(* IEC 61131-3 sources: Masterarbeit/sigmatek/lasalclass2/PW022_virtualization/Network/HW_Network, 1 file *)

(* ---- ONE_HW_Network_Table.st ---- *)
#define OBJECTS_CONFIG

//Define part of class Varan_Base
#ifndef _T_VARANBASE_H
#define _T_VARANBASE_H

#define	VARAN_PLL_OFFSET		16#0140
#define VARAN_MULTIPLE_OFFSET	16#01AC

// version of serial number validation (16#10 = 1.0)
#define SERNO_VALIDATION_VERSION 16#10

#define IsTransparent_IS_AVAILABLE

// Defines for Mutex Generation
#define VARAN_STR_MUTEX_NAME_SEPERATOR ".."
#define VARAN_MUTEX_NAME_END_LENGTH 5
#define VARAN_MUTEX_NAME_MAX_LENGTH 32

#define VARAN_SPI_IDENT_LICENCENO_OFFSET    16#14
#define VARAN_SPI_IDENT_HARDWAREVER_OFFSET  16#18

#endif // _T_VARANBASE_H
#include "..\..\Class\HwControl\HwControl.h"
#include "..\..\Source\interfaces\lsl_st_hardwaretree.h"
//Define part of class BusInterfaceVARAN
#define BUSIF_VARAN_MAX_NR_DO     100
#define BUSIF_VARAN_MAX_NR_MOVEDO 100

#define BUSIF_VARAN_MAX_SDO 1

#define BUSIF_VARAN_BUS_READY_VER 16#1109
#include "..\..\Source\BusInterface.h"
#include "..\..\Source\interfaces\lsl_st_mt.h"
#include "..\..\Source\interfaces\lsl_st_pci.h"
#include "..\..\Class\HwControl\watchdog.h"
#include "..\..\Source\interfaces\lsl_st_sysinfo.h"
#include "..\..\Source\interfaces\lsl_st_systrace.h"
#include "..\..\Class\HwControl\_HWKScope.h"
#include <.\lsl_st_mt.h>
//Define part of class SdiasBase
//Address to access the Dataobject list via SPI SDO Read
#define SDIAS_SPI_DATA_OBJECT_LIST_PAGE_ADDRESS               16#FFFF
#define SDIAS_SPI_DATA_OBJECT_LIST_PAGE_OFFSET                16#00
#define SDIAS_SPI_DATA_OBJECT_LIST_IDENTIFIER                 16#12345678

//Defines the number of optional list elements in the SPI List

#define SDIAS_SPI_NUMBER_OF_OPTIONAL_ELEMENTS                 16

#define SDIAS_SPI_HEADER_BEFORE_OPTIONAL_ELEMENTS             16#18
#define SDIAS_SPI_HARDWARE_VERSION_OFFSET                     16#C
#define SDIAS_SPI_VENDOR_ID_OFFSET                            16#0

#define SDIAS_SPI_MASTER_ADRESS_TRANSMIT_BUFFER0              16#0000
#define SDIAS_SPI_MASTER_ADRESS_TRANSMIT_BUFFER1              16#0080
#define SDIAS_SPI_MASTER_ADRESS_RECEIVE_BUFFER0               16#0000
#define SDIAS_SPI_MASTER_ADRESS_RECEIVE_BUFFER1               16#0080
#define SDIAS_SPI_MASTER_ADRESS_PAGE_ADRESS                   16#0100
#define SDIAS_SPI_MASTER_ADRESS_PREDEFINED_COMMAND_REGISTER   16#0102
#define SDIAS_SPI_MASTER_ADRESS_SINGLE_COMMAND_REGISTER       16#0103
#define SDIAS_SPI_MASTER_ADRESS_STATUS_REGISTER               16#0104
#define SDIAS_SPI_MASTER_ADRESS_REQUEST_REGISTER              16#0105
#define SDIAS_SPI_MASTER_ADRESS_GRANT_REGISTER                16#0106
#define SDIAS_SPI_MASTER_ADRESS_CLEAR_REQUEST_REGISTER        16#0107
#define SDIAS_SPI_MASTER_ADRESS_FEATURE_REGISTER              16#0108

#define SDIAS_SPI_MASTER_SOFTWARE_REQUEST                     1

#define SDIAS_SPI_MASTER_COMMAND_PAGE_READ                    16#01
#define SDIAS_SPI_MASTER_COMMAND_PAGE_PROGRAM                 16#02
#define SDIAS_SPI_MASTER_COMMAND_SECTOR_ERASE                 16#03
#define SDIAS_SPI_MASTER_COMMAND_REBOOT_FPGA                  16#F0

#define SDIAS_SPI_MASTER_STATE_BUSY                           16#00
#define SDIAS_SPI_MASTER_STATE_READY                          16#01

#define SDIAS_SPI_SECTOR_SIZE                                 65536 // 256*256
#define SDIAS_SPI_PAGE_SIZE                                   256

#define SDIAS_SPI_WRITE_MAX_RETRIES                           2
#define SDIAS_SPI_TIMEOUT                                     500  //timeout for spi accesses
#define SDIAS_SPI_LOCK_TIMEOUT                                6   //this value is multiplied with the buscycletime [µs] (6*1000=6.000 msec timeout)

//SPI List IDs
#define SDIAS_SPI_IDENTIFICATION_LIST_ID  1
#define SDIAS_SPI_FLASH_CONFIGURATION_ID  2
#define SDIAS_SPI_VENDOR_NAME_ID          3
#define SDIAS_SPI_DEVICE_NAME_ID          4
#define SDIAS_SPI_SERIAL_NUMBER_ID        5
#define SDIAS_SPI_ORDERING_NUMBER_ID      6
#define SDIAS_SPI_DOCUMENTATION_PDF_ID    7
#define SDIAS_SPI_CALIB_DATA_ID           10
#define SDIAS_SPI_PDO_INFORMATION_ID      128

//SPI Access
#define SDIAS_SPI_ACCESS_ID_HW_TREE          1
#define SDIAS_SPI_ACCESS_ID_HWK_INTERNAL     2
#include "..\..\Class\SdiasManager\SdiasManager.h"
#include "..\..\Class\SdiasBase\SdiasBase.h"
//Define part of class PW022
#define DEVICE_ID_PW022                     1089
// address offsets for SDO communication
#define PW022_ADDR_CFG_MODUL                16#004
// timeouts
#define PW022_SDO_RESPONSE_TIMEOUT          SDIAS_SDO_TIMEOUT * 2
#define PW022_MIN_PERIODE_TIME              100  //minimal allowed periode time * 500nsec
#define PW022_MAX_PERCENT                 10000  //maximal value for percent (100.00)
//Define part of class SafetyUDP
#define SAFETY_UDP_MAX_SOCKETS                6     // Max number of socket

#define SAFETY_UDP_CLT_SEND_OK                0    // Send ok
#define SAFETY_UDP_CLT_INVALID_HANDLE        -1    // Invalid handle
#define SAFETY_UDP_CLT_NOT_OPEN              -2    // Socket is not open
#define SAFETY_UDP_CLT_SEND_FAILED           -3    // Send failed
#define SAFETY_UDP_CLT_SEND_BUFFER_FULL      -4    // Send buffer is full
#define SAFETY_UDP_CLT_DATA_TO_BIG           -5    // Data to big

#define SAFETY_UDP_MAXIMUM_SEGMENT_SIZE    1452    // Maximum of user data

#define SAFETY_UDP_TIMEOUT_OPENSOCKET    (1000)    //timeout for opening socket

#define SAFETY_UDP_RECEIVE_TIMEOUT          800

#define SAFETY_UDP_TX_BUFFER_SIZE          1024
//Define part of class SafetyManager
#define LogBufferSize 1000
#include "..\..\Class\SafetyManager\SafetyManager.h"
#include "..\..\Source\interfaces\lsl_st_safetydll.h"
//Define part of class SdiasManager
#define SDIAS_SDO_MAX_LENGTH              128
#define SDIAS_SDO_RINGBUFFER_NO            64
#define SDIAS_SDO_CHANNEL_NO                3   // fixed in the VI hardware to be 3

// watchdog trigger interval (after 130ms of no trigger the SDIAS HW goes into reset again and takes at least another 10ms to be ready again)
#define SDIAS_WATCHDOG_TRIGGER_TIME        40

// time needed by sdias modules to start up after the watchdog is triggered the first time in ms
#define SDIAS_HARDWARE_STARTUP_TIME        15

// sdias manager needs 2 ticks to handle event for read task (measure sync time)
#define SDIAS_SYNC_MEASURE_TICKS            2

// after activating the PLL SyncOut it takes 3 cycles until the SDIAS sync can be injected
#define SDIAS_CYCLES_WAIT_AFTER_SYNC_ENABLE 3

// wait 1 bus cycle at start to get valid numbers in the task info
#define SDIAS_TASKINFO_READY_TICKS          1

// time to wait (in ms) until other tasks in the same or lower priority than post init have done their stuff
#define SDIAS_WAIT_TIME_IN_POST_INIT        1

#define SIZE_PER_SDIAS_CLIENT               16#0400

// for far memory accesses: 1 module can hold maximum 256 1K blocks (0-255)
#define SDIAS_1K_BLOCK_NO                       256

// far memory accesses maximum length in bytes
#define SDIAS_MAX_SIZE_FAR_MEM_ACCESS           127

#define SDIAS_OFFSET_HW_CONFIG              16#FF00
#define SDIAS_OFFSET_TASK_EVENT_IDS         16#FF10
#define SDIAS_OFFSET_FEATURE_INFO           16#FF18
#define SDIAS_OFFSET_APPLI_LED_STATES       16#FF20
#define SDIAS_OFFSET_SYNC_INJECTION_CFG     16#FF3D
#define SDIAS_OFFSET_TRIGGER_UNIT_SETUP_0   16#FF41
#define SDIAS_OFFSET_TRIGGER_UNIT_SETUP_1   16#FF45
#define SDIAS_OFFSET_TASK_START_CFG_0       16#FF60
#define SDIAS_OFFSET_TASK_CONFIG_0          16#FF86
#define SDIAS_OFFSET_TASK_CONFIG_1          16#FF96
#define SDIAS_OFFSET_TASK_INFO_1            16#FF94
#define SDIAS_OFFSET_TASK_HANDSHAKE_1       16#FF9B
#define SDIAS_OFFSET_TASK_DURATION_TIME_1   16#FF9C
#define SDIAS_OFFSET_TASK_DURATION_TIME_2   16#FFAC
#define SDIAS_OFFSET_TASK_CONFIG_2          16#FFA6

#define SDIAS_RETRIES_ALLOWED         2

// mask to get global error flag out of message counter byte of SDO responses
#define SDIAS_MASK_GLOBAL_ERROR_FLAG        16#80

// mask to get message counter out of message counter byte of SDO responses
#define SDIAS_MASK_MESSAGE_COUNTER          16#3F

#define SDIAS_EVENT_MASK_ID_SYNC_OUT0       16#10
#define SDIAS_EVENT_MASK_ID_SYNC_OUT1       16#11
#define SDIAS_EVENT_MASK_ID_SYNC_OUT2       16#12
#define SDIAS_EVENT_MASK_ID_SYNC_OUT3       16#13

#define SDIAS_MANAGER_SYNC_SYNCOUT_ID       16#85
#define SDIAS_TASK_START_EVENT_SYNCOUT_ID   16#86

#define SDIAS_PLACE_NO_MODULE_ADDED_SO_FAR  16#80000000

#define SDIAS_TRIGGER_UNIT_BYTE_SIZE        2

#define SDIAS_WAIT_TIME_FIRMWARE_HANDSHAKE  5 * 1000

// if the firmware version is below this, there might be problems with SCP111 and other modules => print warning at startup
#define SDIAS_FW_VERSION_SDO_ERROR_FIXED    16#120

// if the protocol version ist below this, Control Read/Broadcast Write Command is not supported by sdiasmanager
#define SDIAS_PROTOCOLVERSION_BROADCAST     16#120

// if the cil version ist below this, Control Read/Broadcast Write Command is not supported by OS for local SDIAS.
#define SDIAS_CILVERSION_BROADCAST         16#5001

// timeout for blocking the init during initialisation (in ms)
#define SDIAS_INIT_BLOCK_TIMEOUT            20 * 1000

#define SDIAS_MUTEX_NAME_END_LENGTH 3
#define SDIAS_MUTEX_NAME_MAX_LENGTH 32
#define SDIAS_MUTEX_STR_SEPERATOR   ".."

//#define SDIAS_RT_TIME_MEASUREMENT
#ifdef SDIAS_RT_TIME_MEASUREMENT
  #pragma message("ATTENTION: SDIAS real time measurement is active and needs additional ressources in the realtime task")
#endif

(* SDIAS data object commands  *)
#define	 SDIAS_CMD_END							  0x00			(* End command										          *)
#define	 SDIAS_CMD_ACC_MEMORY				  0x01			(* Access dpram memory								      *)
#define	 SDIAS_CMD_ACC_CONTROL				0x02			(* Access dpram control memory						  *)
#define	 SDIAS_CMD_GLOBAL						  0x03			(* SDIAS global command								      *)
#define	 SDIAS_CMD_COPY_LOCAL					0x04			(* DPRAM copy command in local dpram				*)
#define	 SDIAS_CMD_JMP_LOCAL					0x05			(* DPRAM jump command in local dpram 				*)
#define  SDIAS_CMD_ACC_MEMORY_FAR     0x07      (* SDIAS Far Memory Access                  *)

(* SDIAS defines for data object handling *)
// Write data oject list
#define	 SDIAS_DOL_WRITE_USAGE_DOL_EMPTY	  0x20			(* Usage of empty write dol list (wachtdog trigger + end command)   *)
#define	 SDIAS_DOL_WRITE_USAGE_DTA_EMPTY	  0x03			(* Usage of empty write dol data (DO ctrl of 2x copy command for task information + DO ctrl of watchdog trigger      *)
#define	 SDIAS_DOL_WRITE_OFFSET_END_CMD			0x10			(* One data object in list - offset = 1 DO size = 0x10						  *)
#define	 SDIAS_DOL_WRITE_OFFSET_FIRST_DTA		0x02			(* Offset of first data byte of second copy command = 2 (DO ctrl)   *)
#define	 SDIAS_DOL_WRITE_OFFSET_LAST_DTA		0x02			(* Offset of last data byte of second copy command = 2 (DO ctrl )   *)

// Read data oject list
#define	 SDIAS_DOL_READ_USAGE_DOL_EMPTY	    0x30			(* Usage of empty read dol list (2x task info copy command + end command)   *)
#define	 SDIAS_DOL_READ_USAGE_DTA_EMPTY	    0x0D			(* Usage of empty write dol data (DO ctrl of 2x copy command for task information + DO ctrl of watchdog trigger      *)
#define	 SDIAS_DOL_READ_OFFSET_END_CMD			0x20			(* One data object in list - offset = 1 DO size = 0x10						          *)
#define	 SDIAS_DOL_READ_OFFSET_FIRST_DTA		0x07			(* Offset of first data byte of second copy command = 7 = DO state          *)
#define	 SDIAS_DOL_READ_OFFSET_LAST_DTA		  0x0C			(* Offset of last data byte of second copy command = 12 (last byte of task information)       *)

//Versionsnumber where SDIAS SPI Read Accesses are available
#define  SDIAS_SDO_SPI_FIRMWARE_VERSION_AVAILABLE 16#0120

//error info mask
#define  SDIAS_ERROR_INFO_MASK    2#1000011000011111

// Broadcast DO Info
#define SDIAS_OFFSET_CLIENT_CTRLTIMESTAMP   16#0190
#define SDIAS_NR_TIMEBROADCAST_DOS 2
#define SDIAS_TIMEBROADCAST_SUBCMD 16#B0
#include "..\..\source\interfaces\lsl_st_pll.h"
//Define part of class VaranManager
#define SIZE_PAYLOAD_FRAME_HEADER_DO      16#38  // Const because datasize is in the Payload DOs
#define SIZE_PAYLOAD_IRQ_FRAME_HEADER_DO  16#40  // Const because datasize is in the Payload DOs

#define VM_MAX_POST_INIT_MODULES  1000

#define VM_OBJECT_PATH            16#81000002   // Object Path for Varanmanager Length = 2 (First 2byte), Domain = 0 (3rd byte), Escape Sequence Varan (4th byte)
#include "..\..\Class\VaranManager\VaranManager.h"
#include "..\..\Source\interfaces\lsl_st_kernel.h"
//Define part of class VaranManager_2
// needed to use the same code as the other managing modules
#define VM2_SYNCHRON SuperiorSystemOK

#define VM2_SDO_INIT_CMD_LENGTH   12
//Define part of class VI021
#define DEVICE_ID_VI022 1233

FUNCTION GLOBAL TAB ONE_HW_Network
-1$UINT, 0$UINT,
0$UINT, 0$UINT,

26$UDINT,
TO_UDINT(2897291062), "ASCII_BIN", 1$UINT, 21$UINT, 1$UINT,
TO_UDINT(24783181), "BusInterfaceVARAN", 1$UINT, 75$UINT, 0$UINT,
TO_UDINT(794617671), "CriticalSection", 0$UINT, 4$UINT, 2$UINT,
TO_UDINT(3238133653), "Hub_Base", 1$UINT, 21$UINT, 1$UINT,
TO_UDINT(1770276445), "Hub_Base_Root", 2$UINT, 11$UINT, 2$UINT,
TO_UDINT(3078259981), "HwcLogging", 1$UINT, 0$UINT, 1$UINT,
TO_UDINT(2471641665), "HwControl", 5$UINT, 21$UINT, 1$UINT,
TO_UDINT(1193052171), "HwControlBase", 1$UINT, 10$UINT, 0$UINT,
TO_UDINT(4260294091), "HWRtPostScan", 1$UINT, 0$UINT, 1$UINT,
TO_UDINT(2225119864), "MerkerEx", 1$UINT, 22$UINT, 4$UINT,
TO_UDINT(2837966764), "PW022", 1$UINT, 5$UINT, 3$UINT,
TO_UDINT(3591333481), "RamFile", 1$UINT, 9$UINT, 1$UINT,
TO_UDINT(1799751072), "SafetyManager", 2$UINT, 26$UINT, 1$UINT,
TO_UDINT(3727715967), "SafetyUDP", 1$UINT, 4$UINT, 0$UINT,
TO_UDINT(3175101883), "SdiasBase", 1$UINT, 60$UINT, 0$UINT,
TO_UDINT(4173303375), "SdiasHubBase", 1$UINT, 10$UINT, 1$UINT,
TO_UDINT(2118381352), "SdiasManager", 1$UINT, 97$UINT, 1$UINT,
TO_UDINT(736632136), "Steuerung", 0$UINT, 0$UINT, 1$UINT,
TO_UDINT(1850111279), "String", 1$UINT, 11$UINT, 4$UINT,
TO_UDINT(2898603620), "StringInternal", 1$UINT, 85$UINT, 0$UINT,
TO_UDINT(862125188), "Varan_Base", 2$UINT, 20$UINT, 0$UINT,
TO_UDINT(2940693151), "VaranManager", 3$UINT, 7$UINT, 0$UINT,
TO_UDINT(4019434288), "VaranManager_2", 2$UINT, 9$UINT, 1$UINT,
TO_UDINT(4035182347), "VaranManager_Base", 1$UINT, 26$UINT, 0$UINT,
TO_UDINT(262695706), "VI021", 1$UINT, 101$UINT, 1$UINT,
TO_UDINT(3232495061), "VirtualBaseInit", 1$UINT, 3$UINT, 0$UINT,

1$UINT, TO_UDINT(1973273396), "VARANMANAGER_21\_BASE\ASCII_BIN1",

1$UINT, TO_UDINT(2972590922), "HWCONTROL1\SAFETYMANAGER\UDPRECEIVEDATA",
1$UINT, TO_UDINT(1868223583), "HWCONTROL1\SAFETYMANAGER\UDPSENDDATA",

1$UINT, TO_UDINT(658018123), "VI0211\HUB_BASE1",

1$UINT, TO_UDINT(980975553), "VARANMANAGER_21\HUB_BASE_ROOT0",
1$UINT, TO_UDINT(1300189015), "VARANMANAGER_21\HUB_BASE_ROOT1",

1$UINT, TO_UDINT(3105254819), "HWCONTROL1\HWCLOGGING",

_NO_ATTR, TO_UDINT(2190789875), "HWCONTROL1",

1$UINT, TO_UDINT(1673205898), "HWCONTROL1\HWRTPOSTSCAN",

1$UINT, TO_UDINT(2963574667), "PW022_1\_BASE\SERIALNOSTR\MERKEREX0",
1$UINT, TO_UDINT(1616831850), "PW022_1_COPY\_BASE\SERIALNOSTR\MERKEREX0",
1$UINT, TO_UDINT(404369275), "PW022_1_COPY_COPY\_BASE\SERIALNOSTR\MERKEREX0",
1$UINT, TO_UDINT(1965133148), "VI0211\_BASE\_BASE\SERIALNOSTR\MERKEREX0",

_NO_ATTR, TO_UDINT(522450549), "PW022_1",
_NO_ATTR, TO_UDINT(1130690254), "PW022_1_COPY",
_NO_ATTR, TO_UDINT(1202210518), "PW022_1_COPY_COPY",

1$UINT, TO_UDINT(4171808520), "VI0211\_BASE\_BASE\SERNOBACKUP",

1$UINT, TO_UDINT(1778590035), "HWCONTROL1\SAFETYMANAGER",

1$UINT, TO_UDINT(1199943557), "VI0211\SDIASHUBBASE",

1$UINT, TO_UDINT(3245985506), "VI0211\SDIASMANAGER",

_NO_ATTR, TO_UDINT(4226862600), "STEUERUNG1",

1$UINT, TO_UDINT(2032061554), "PW022_1\_BASE\SERIALNOSTR",
1$UINT, TO_UDINT(1101856492), "PW022_1_COPY\_BASE\SERIALNOSTR",
1$UINT, TO_UDINT(2768093490), "PW022_1_COPY_COPY\_BASE\SERIALNOSTR",
1$UINT, TO_UDINT(3053332208), "VI0211\_BASE\_BASE\SERIALNOSTR",

_NO_ATTR, TO_UDINT(2783595688), "VARANMANAGER_21",

_NO_ATTR, TO_UDINT(2125577894), "VI0211",

//Internal connections
0$UDINT,
20$UDINT,
TO_UDINT(7), "SafetyManager", TO_UDINT(17),
TO_UDINT(7), "HWRtPostScan", TO_UDINT(8),
TO_UDINT(7), "HwcLogging", TO_UDINT(6),
TO_UDINT(13), "SerialNoStr", TO_UDINT(21),
TO_UDINT(14), "SerialNoStr", TO_UDINT(22),
TO_UDINT(15), "SerialNoStr", TO_UDINT(23),
TO_UDINT(17), "UdpSendData", TO_UDINT(2),
TO_UDINT(17), "UdpReceiveData", TO_UDINT(1),
TO_UDINT(21), "MerkerEx0", TO_UDINT(9),
TO_UDINT(22), "MerkerEx0", TO_UDINT(10),
TO_UDINT(23), "MerkerEx0", TO_UDINT(11),
TO_UDINT(24), "MerkerEx0", TO_UDINT(12),
TO_UDINT(25), "ASCII_BIN1", TO_UDINT(0),
TO_UDINT(25), "Hub_Base_Root0", TO_UDINT(4),
TO_UDINT(25), "Hub_Base_Root1", TO_UDINT(5),
TO_UDINT(26), "SerialNoStr", TO_UDINT(24),
TO_UDINT(26), "SerNoBackup", TO_UDINT(16),
TO_UDINT(26), "Hub_Base1", TO_UDINT(3),
TO_UDINT(26), "SdiasManager", TO_UDINT(19),
TO_UDINT(26), "SdiasHubBase", TO_UDINT(18),
0$UDINT,
28$UDINT,
TO_UDINT(3), "VaranIn", TO_UDINT(26), "State",
TO_UDINT(4), "VaranConnect", TO_UDINT(25), "Control",
TO_UDINT(5), "VaranConnect", TO_UDINT(25), "Control",
TO_UDINT(8), "toHwControlBase", TO_UDINT(7), "Control",
TO_UDINT(13), "SdiasIn", TO_UDINT(18), "ClassSvr",
TO_UDINT(14), "SdiasIn", TO_UDINT(18), "ClassSvr",
TO_UDINT(15), "SdiasIn", TO_UDINT(18), "ClassSvr",
TO_UDINT(17), "To_HwControl", TO_UDINT(7), "Control",
TO_UDINT(18), "ToNextSDIAS", TO_UDINT(19), "ClassState",
TO_UDINT(19), "ToBusInterface", TO_UDINT(26), "CallCommand",
TO_UDINT(20), "cPeriodeDuration_ch1", TO_UDINT(13), "PeriodeDuration_Ch1",
TO_UDINT(20), "cPWMOnTime_ch1", TO_UDINT(13), "PWMOnTime_Ch1",
TO_UDINT(20), "cPeriodeDuration_ch2", TO_UDINT(13), "PeriodeDuration_Ch2",
TO_UDINT(20), "cPWMOnTime_ch2", TO_UDINT(13), "PWMOnTime_Ch2",
TO_UDINT(20), "cPeriodeDuration_ch3", TO_UDINT(14), "PeriodeDuration_Ch1",
TO_UDINT(20), "cPWMOnTime_ch3", TO_UDINT(14), "PWMOnTime_Ch1",
TO_UDINT(20), "cPeriodeDuration_ch4", TO_UDINT(14), "PeriodeDuration_Ch2",
TO_UDINT(20), "cPWMOnTime_ch4", TO_UDINT(14), "PWMOnTime_Ch2",
TO_UDINT(20), "cPeriodeDuration_ch5", TO_UDINT(15), "PeriodeDuration_Ch1",
TO_UDINT(20), "cPWMOnTime_ch5", TO_UDINT(15), "PWMOnTime_Ch1",
TO_UDINT(20), "cPeriodeDuration_ch6", TO_UDINT(15), "PeriodeDuration_Ch2",
TO_UDINT(20), "cPWMOnTime_ch6", TO_UDINT(15), "PWMOnTime_Ch2",
TO_UDINT(21), "DataBuffer", TO_UDINT(9), "m_udLength",
TO_UDINT(22), "DataBuffer", TO_UDINT(10), "m_udLength",
TO_UDINT(23), "DataBuffer", TO_UDINT(11), "m_udLength",
TO_UDINT(24), "DataBuffer", TO_UDINT(12), "m_udLength",
TO_UDINT(25), "To_HwControl", TO_UDINT(7), "Control",
TO_UDINT(26), "VaranIn", TO_UDINT(4), "Control",

//Initialization values
0$UDINT,
49$UDINT,
TO_UDINT(3), "Splitter_Place", TO_UDINT(0),//|HW_Network.VI0211\Hub_Base1.Splitter_Place;
TO_UDINT(4), "Splitter_Place", TO_UDINT(0),//|HW_Network.VaranManager_21\Hub_Base_Root0.Splitter_Place;
TO_UDINT(5), "Splitter_Place", TO_UDINT(1),//|HW_Network.VaranManager_21\Hub_Base_Root1.Splitter_Place;
TO_UDINT(7), "UdpSafetyPort", TO_UDINT(10823),//|HW_Network.HwControl1.UdpSafetyPort;
TO_UDINT(7), "InterfaceNo", TO_UDINT(1),//|HW_Network.HwControl1.InterfaceNo;
TO_UDINT(7), "RtTaskSync", TO_UDINT(0),//|HW_Network.HwControl1.RtTaskSync;
TO_UDINT(9), "ThreadSafe", TO_UDINT(0),//|HW_Network.SerialNoStr\_base\PW022_1\MerkerEx0.ThreadSafe;
TO_UDINT(10), "ThreadSafe", TO_UDINT(0),//|HW_Network.SerialNoStr\_base\PW022_1_Copy\MerkerEx0.ThreadSafe;
TO_UDINT(11), "ThreadSafe", TO_UDINT(0),//|HW_Network.SerialNoStr\_base\PW022_1_Copy_Copy\MerkerEx0.ThreadSafe;
TO_UDINT(12), "ThreadSafe", TO_UDINT(0),//|HW_Network.SerialNoStr\_base\_base\VI0211\MerkerEx0.ThreadSafe;
TO_UDINT(13), "LEDControl", TO_UDINT(0),//|HW_Network.PW022_1.LEDControl;
TO_UDINT(13), "PeriodeDuration_Ch1", TO_UDINT(100),//|HW_Network.PW022_1.PeriodeDuration_Ch1;
TO_UDINT(13), "PeriodeDuration_Ch2", TO_UDINT(100),//|HW_Network.PW022_1.PeriodeDuration_Ch2;
TO_UDINT(13), "Place", TO_UDINT(0),//|HW_Network.PW022_1.Place;
TO_UDINT(13), "Required", TO_UDINT(1),//|HW_Network.PW022_1.Required;
TO_UDINT(13), "PWMUnitMode", TO_UDINT(0),//|HW_Network.PW022_1.PWMUnitMode;
TO_UDINT(14), "LEDControl", TO_UDINT(0),//|HW_Network.PW022_1_Copy.LEDControl;
TO_UDINT(14), "PeriodeDuration_Ch1", TO_UDINT(100),//|HW_Network.PW022_1_Copy.PeriodeDuration_Ch1;
TO_UDINT(14), "PeriodeDuration_Ch2", TO_UDINT(100),//|HW_Network.PW022_1_Copy.PeriodeDuration_Ch2;
TO_UDINT(14), "Place", TO_UDINT(1),//|HW_Network.PW022_1_Copy.Place;
TO_UDINT(14), "Required", TO_UDINT(0),//|HW_Network.PW022_1_Copy.Required;
TO_UDINT(14), "PWMUnitMode", TO_UDINT(0),//|HW_Network.PW022_1_Copy.PWMUnitMode;
TO_UDINT(15), "LEDControl", TO_UDINT(0),//|HW_Network.PW022_1_Copy_Copy.LEDControl;
TO_UDINT(15), "PeriodeDuration_Ch1", TO_UDINT(100),//|HW_Network.PW022_1_Copy_Copy.PeriodeDuration_Ch1;
TO_UDINT(15), "PeriodeDuration_Ch2", TO_UDINT(100),//|HW_Network.PW022_1_Copy_Copy.PeriodeDuration_Ch2;
TO_UDINT(15), "Place", TO_UDINT(2),//|HW_Network.PW022_1_Copy_Copy.Place;
TO_UDINT(15), "Required", TO_UDINT(0),//|HW_Network.PW022_1_Copy_Copy.Required;
TO_UDINT(15), "PWMUnitMode", TO_UDINT(0),//|HW_Network.PW022_1_Copy_Copy.PWMUnitMode;
TO_UDINT(16), "Setup", TO_UDINT(2#1101),//|HW_Network._base\_base\VI0211\SerNoBackup.Setup;
TO_UDINT(17), "UdpSafetyPort", TO_UDINT(10823),//|HW_Network.HwControl1\SafetyManager.UdpSafetyPort;
TO_UDINT(17), "InterfaceNo", TO_UDINT(1),//|HW_Network.HwControl1\SafetyManager.InterfaceNo;
TO_UDINT(17), "UdpSafetyRequestCycle", TO_UDINT(UDP_MIN_REQUEST_TIME),//|HW_Network.HwControl1\SafetyManager.UdpSafetyRequestCycle;
TO_UDINT(17), "UdpSafetyResponseTimeout", TO_UDINT(UDP_MIN_RESPONSE_TIMEOUT),//|HW_Network.HwControl1\SafetyManager.UdpSafetyResponseTimeout;
TO_UDINT(18), "SplitterPlace", TO_UDINT(0),//|HW_Network.VI0211\SdiasHubBase.SplitterPlace;
TO_UDINT(19), "DeviceID", TO_UDINT(1187),//|HW_Network.VI0211\SdiasManager.DeviceID;
TO_UDINT(19), "AutoFarMem", TO_UDINT(0),//|HW_Network.VI0211\SdiasManager.AutoFarMem;
TO_UDINT(21), "SingleRealloc", TO_UDINT(1),//|HW_Network._base\PW022_1\SerialNoStr.SingleRealloc;
TO_UDINT(22), "SingleRealloc", TO_UDINT(1),//|HW_Network._base\PW022_1_Copy\SerialNoStr.SingleRealloc;
TO_UDINT(23), "SingleRealloc", TO_UDINT(1),//|HW_Network._base\PW022_1_Copy_Copy\SerialNoStr.SingleRealloc;
TO_UDINT(24), "SingleRealloc", TO_UDINT(1),//|HW_Network._base\_base\VI0211\SerialNoStr.SingleRealloc;
TO_UDINT(25), "VaranManagerTime", TO_UDINT(10000000),//|HW_Network.VaranManager_21.VaranManagerTime;
TO_UDINT(25), "VaranManagerNr", TO_UDINT(0),//|HW_Network.VaranManager_21.VaranManagerNr;
TO_UDINT(25), "PayloadFrame", TO_UDINT(2),//|HW_Network.VaranManager_21.PayloadFrame;
TO_UDINT(25), "CoreSelect", TO_UDINT(0),//|HW_Network.VaranManager_21.CoreSelect;
TO_UDINT(25), "InterframeGap", TO_UDINT(0),//|HW_Network.VaranManager_21.InterframeGap;
TO_UDINT(26), "Required", TO_UDINT(1),//|HW_Network.VI0211.Required;
TO_UDINT(26), "Transparent", TO_UDINT(0),//|HW_Network.VI0211.Transparent;
TO_UDINT(26), "TimeBase", TO_UDINT(0),//|HW_Network.VI0211.TimeBase;
TO_UDINT(26), "TimeBaseOffset", TO_UDINT(0),//|HW_Network.VI0211.TimeBaseOffset;

//Symbolic initialization values
0$UDINT,
0$UDINT,

//Initialization of string values
0$UDINT,
0$UDINT,

//Configuration of tasks (RealTime, Cyclic, Background)
0$UDINT,
2$UDINT,
TO_UDINT(20), (1)$UDINT, 4194303$DINT, 	//STEUERUNG1
TO_UDINT(8), (1)$UDINT, 4194304$DINT, 	//HWCONTROL1\HWRTPOSTSCAN

0$UDINT,
0$UDINT,

0$UDINT,
0$UDINT,

//External connections
0$UDINT,
0$UDINT,

//Magic internal connections
0$UDINT,
3$UDINT,
TO_UDINT(17), "UdpSafetyPort", TO_UDINT(7), "UdpSafetyPort",
TO_UDINT(17), "InterfaceNo", TO_UDINT(7), "InterfaceNo",
TO_UDINT(17), "SafetyDomainTimeout", TO_UDINT(7), "SafetyDomainTimeout",

//Configuration of timeslots of tasks (RealTime, Cyclic)
#ifdef __LSLLDR_TIMESLOTS__
0$UDINT,
0$UDINT,

0$UDINT,
0$UDINT,

#endif //__LSLLDR_TIMESLOTS__

//MultiMaster connections
#ifdef __LSLLDR_MULTIMASTER__
0$UDINT,
0$UDINT,
#endif //__LSLLDR_MULTIMASTER__

//Configuration for task ID (RealTime, CyclicTime)
#ifdef __LSLLDR_TASKID__
"\\\\TASKS2  "
0$UDINT,
2$UDINT,
(0)$UDINT, 	//STEUERUNG1
(0)$UDINT, 	//HWCONTROL1\HWRTPOSTSCAN

0$UDINT,
0$UDINT,

0$UDINT,
0$UDINT,

#endif //__LSLLDR_TASKID__

END_FUNCTION
